(* IEC 61131-3 sources: rusty/tests/lit/single/variadics, 4 files *)

(* ---- bitaccess_xor_printf.st ---- *)
// RUN: %COMPILE %s && %RUN | %CHECK %s
// Verifies that a boolean XOR expression involving a direct bit-access is
// correctly promoted to i32 when passed as a variadic argument.
// Without the promotion the i1 result can be clobbered by the subsequent MUX
// call, causing the same expression to print different values before and after.

FUNCTION foo
    VAR
        vTrue  : BOOL := TRUE;
        vFalse : BOOL := FALSE;
        arrLword : LWORD := 16#abcdefabcdefabcd;
        // bit 27 of arrLword = 1, so:
        //   bit27 XOR TRUE  = 0
        //   bit27 XOR FALSE = 1
    END_VAR

    // Simplified bit-access via %x27 (same as %d0.%w1.%B1.%x3)
    printf('before mux xor TRUE: %u$N', arrLword.%x27 XOR vTrue);   // CHECK: before mux xor TRUE: 0
    MUX(0, 255, 255);
    printf('after mux xor TRUE: %u$N',  arrLword.%x27 XOR vTrue);   // CHECK: after mux xor TRUE: 0

    printf('before mux xor FALSE: %u$N', arrLword.%x27 XOR vFalse); // CHECK: before mux xor FALSE: 1
    MUX(0, 255, 255);
    printf('after mux xor FALSE: %u$N',  arrLword.%x27 XOR vFalse); // CHECK: after mux xor FALSE: 1

    // Chain-access form from the original bug report
    printf('chain before mux: %u$N', arrLword.%d0.%w1.%B1.%x3 XOR vTrue);  // CHECK: chain before mux: 0
    MUX(0, 255, 255);
    printf('chain after mux: %u$N',  arrLword.%d0.%w1.%B1.%x3 XOR vTrue);  // CHECK: chain after mux: 0

END_FUNCTION

FUNCTION main : DINT
    foo();
END_FUNCTION

(* ---- implicit_types_passed_correctly.st ---- *)
// RUN: %COMPILE %s && %RUN | %CHECK %s
FUNCTION main: DINT
    VAR
        x : UDINT := 21;
        y : LREAL := 42;
    END_VAR

    // CHECK: X(21): Y = 42.000000
    printf('X(%u): Y = %f', x, y);
END_FUNCTION

(* ---- string_passed_as_pointer.st ---- *)
// RUN: %COMPILE %s && %RUN | %CHECK %s
// Test that STRING types are correctly passed as pointers to variadic functions
// per C spec (strings decay to char* pointers)
// CHECK: My string is: hello
FUNCTION main : DINT
VAR
    myString : STRING := 'hello';
END_VAR
    printf('My string is: %s$N', myString);
END_FUNCTION

(* ---- bool_printf.st ---- *)
// RUN: %COMPILE %s && %RUN | %CHECK %s
// Verifies that BOOL values and boolean expressions are correctly promoted to
// 32-bit integers when passed as variadic arguments, matching C default argument
// promotion rules. Without this promotion the values can appear as 255/254 at
// -Onone because the raw i1/i8 is misread by printf.

PROGRAM mainProg
VAR
    vTrue  : BOOL := TRUE;
    vFalse : BOOL := FALSE;
END_VAR

    // Literals
    printf('FALSE: %u$N', FALSE);           // CHECK: FALSE: 0
    printf('TRUE: %u$N', TRUE);             // CHECK: TRUE: 1

    // NOT of literals
    printf('NOT FALSE: %u$N', NOT FALSE);   // CHECK: NOT FALSE: 1
    printf('NOT TRUE: %u$N', NOT TRUE);     // CHECK: NOT TRUE: 0

    // AND expressions
    printf('TRUE AND FALSE: %u$N', TRUE AND FALSE);   // CHECK: TRUE AND FALSE: 0
    printf('TRUE AND TRUE: %u$N', TRUE AND TRUE);     // CHECK: TRUE AND TRUE: 1

    // NOT of AND expressions
    printf('NOT (TRUE AND FALSE): %u$N', NOT (TRUE AND FALSE));  // CHECK: NOT (TRUE AND FALSE): 1
    printf('NOT (TRUE AND TRUE): %u$N', NOT (TRUE AND TRUE));    // CHECK: NOT (TRUE AND TRUE): 0

    // OR expressions
    printf('FALSE OR FALSE: %u$N', FALSE OR FALSE);  // CHECK: FALSE OR FALSE: 0
    printf('TRUE OR FALSE: %u$N', TRUE OR FALSE);    // CHECK: TRUE OR FALSE: 1

    // Variables
    printf('vFalse: %u$N', vFalse);        // CHECK: vFalse: 0
    printf('vTrue: %u$N', vTrue);          // CHECK: vTrue: 1

    // NOT of variables
    printf('NOT vFalse: %u$N', NOT vFalse); // CHECK: NOT vFalse: 1
    printf('NOT vTrue: %u$N', NOT vTrue);   // CHECK: NOT vTrue: 0

    // NOT of variable AND expressions
    printf('NOT (vTrue AND vFalse): %u$N', NOT (vTrue AND vFalse)); // CHECK: NOT (vTrue AND vFalse): 1
    printf('NOT (vTrue AND vTrue): %u$N', NOT (vTrue AND vTrue));   // CHECK: NOT (vTrue AND vTrue): 0

END_PROGRAM

FUNCTION main : DINT
    mainProg();
END_FUNCTION
